Omron CX-Programmer project NewProject (CX-Programmer 9.75)

# PLC wastewater_treatment: CP1E E20

## Global symbols (name address type ; comment)
0.00 BOOL  ; PB_START
0.03 BOOL  ; AUGER_CHECK
0.01 BOOL  ; PB_STOP
0.02 BOOL  ; estop_high
100.00 BOOL  ; AUGER_RUN
100.01 BOOL  ; FLUSH_SOLENOID
100.02 BOOL  ; ACTUATOR_EXTEND
100.03 BOOL  ; ACTUATOR_RETRACT
100.04 BOOL  ; ALARM
90 CHANNEL  ; FLOW<SETPOINT
D10 CHANNEL  ; FLOW
T000 BOOL  ; T_FLOW_DELAY
T001 BOOL  ; T_JAM_RELIEF
T002 BOOL  ; T_PURGE_FLUSH
T003 BOOL  ; T_PRECHOKE
W0.00 BOOL  ; SYS_RUN
W0.01 BOOL  ; SEQ_PRECHOKE
W0.02 BOOL  ; SEQ_DEWATER
W0.03 BOOL  ; JAM_RELIEF
W0.04 BOOL  ; SEQ_SHUTDOWN
W0.05 BOOL  ; ALM_LOW_FLOW

## Program NewProgram1 (cyclic task 0)

### Section Section1

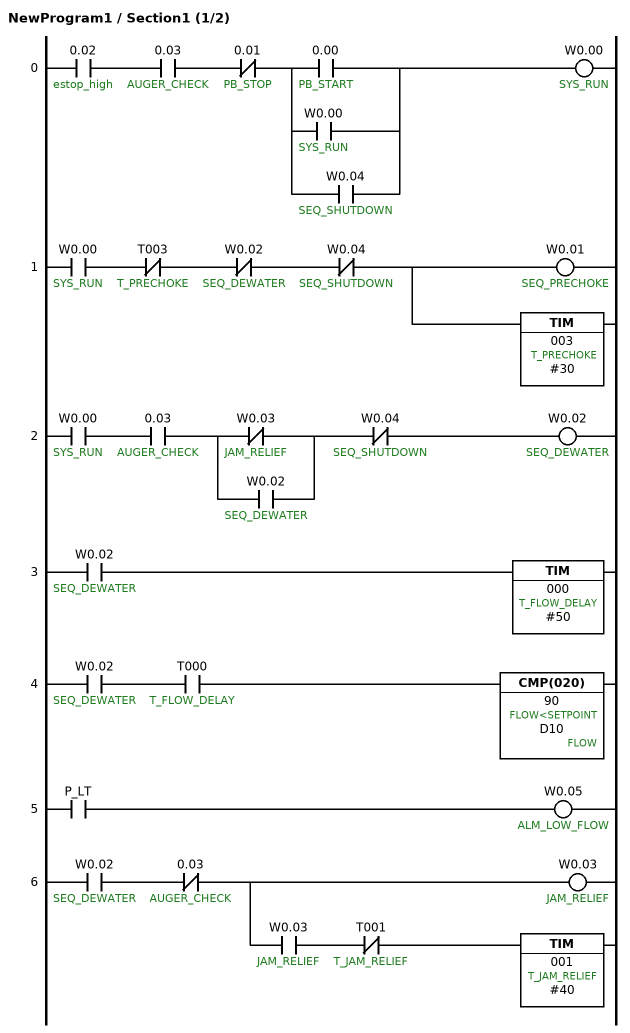
; rung 0
LD 0.02  ; estop_high
AND 0.03  ; AUGER_CHECK
ANDNOT 0.01  ; PB_STOP
LD 0.00  ; PB_START
OR W0.00  ; SYS_RUN
OR W0.04  ; SEQ_SHUTDOWN
ANDLD
OUT W0.00  ; SYS_RUN
; rung 1
LD W0.00  ; SYS_RUN
ANDNOT T003  ; T_PRECHOKE
ANDNOT W0.02  ; SEQ_DEWATER
ANDNOT W0.04  ; SEQ_SHUTDOWN
OUT W0.01  ; SEQ_PRECHOKE
TIM 003 #30  ; T_PRECHOKE
; rung 2
LD W0.00  ; SYS_RUN
AND 0.03  ; AUGER_CHECK
LDNOT W0.03  ; JAM_RELIEF
OR W0.02  ; SEQ_DEWATER
ANDLD
ANDNOT W0.04  ; SEQ_SHUTDOWN
OUT W0.02  ; SEQ_DEWATER
; rung 3
LD W0.02  ; SEQ_DEWATER
TIM 000 #50  ; T_FLOW_DELAY
; rung 4
LD W0.02  ; SEQ_DEWATER
AND T000  ; T_FLOW_DELAY
CMP(020) 90 D10  ; FLOW<SETPOINT, FLOW
; rung 5
LD P_LT
OUT W0.05  ; ALM_LOW_FLOW
; rung 6
LD W0.02  ; SEQ_DEWATER
ANDNOT 0.03  ; AUGER_CHECK
OUT W0.03  ; JAM_RELIEF
AND W0.03  ; JAM_RELIEF
ANDNOT T001  ; T_JAM_RELIEF
TIM 001 #40  ; T_JAM_RELIEF

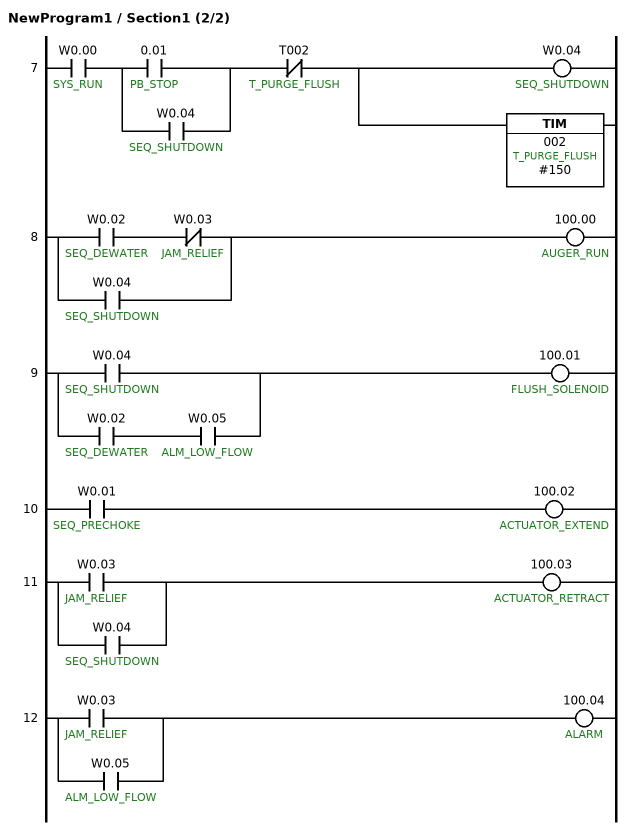
; rung 7
LD W0.00  ; SYS_RUN
LD 0.01  ; PB_STOP
OR W0.04  ; SEQ_SHUTDOWN
ANDLD
ANDNOT T002  ; T_PURGE_FLUSH
OUT W0.04  ; SEQ_SHUTDOWN
TIM 002 #150  ; T_PURGE_FLUSH
; rung 8
LD W0.02  ; SEQ_DEWATER
ANDNOT W0.03  ; JAM_RELIEF
OR W0.04  ; SEQ_SHUTDOWN
OUT 100.00  ; AUGER_RUN
; rung 9
LD W0.04  ; SEQ_SHUTDOWN
LD W0.02  ; SEQ_DEWATER
AND W0.05  ; ALM_LOW_FLOW
ORLD
OUT 100.01  ; FLUSH_SOLENOID
; rung 10
LD W0.01  ; SEQ_PRECHOKE
OUT 100.02  ; ACTUATOR_EXTEND
; rung 11
LD W0.03  ; JAM_RELIEF
OR W0.04  ; SEQ_SHUTDOWN
OUT 100.03  ; ACTUATOR_RETRACT
; rung 12
LD W0.03  ; JAM_RELIEF
OR W0.05  ; ALM_LOW_FLOW
OUT 100.04  ; ALARM

### Section END
; rung 0
END(001)